TYPE ST_NestProcessResult :
STRUCT
	bResultValid        : BOOL;
    bPass               : BOOL;
    bFail               : BOOL;
    bDispositionSent    : BOOL;
END_STRUCT
END_TYPE

(* stored: Version 1.1.0.1
   DUT ST_NestProcessResult: Id {403df8ef-2425-404f-9223-dd5ae33d0d7c} *)
